(* IEC 61131-3 sources: JingjiangArm/moonboxpro_arm_8.4/Application/Application/任务列表/Main_Task/套色调整/套色新算法/PID_GET/Arc_pidh, 3 files *)

(* ---- DOUBLE_INTER.st ---- *)
(*@CES
Name=DOUBLE_INTER
Type=FunctionBlock
TypeGuid=6f9dac99-8de1-4efc-8465-68ac443b7d08
Guid=ffc9ca76-f385-4e76-b007-d8ddf6459d90
HasDeclaration=True
HasImplementation=True
*)
{DECLARATION}
FUNCTION DOUBLE_INTER : LREAL
VAR_INPUT
    (* --- 运行时输入 --- *)
    lrV_m_min   : LREAL;    (* 线速度 (m/min)，需在内部转换为 m/s *)
    lrY_Meas    : LREAL;    (* 测量套色误差 (mm) *)
    bEnable     : BOOL;     (* 控制器使能 *)

    (* --- 配置参数 (PSO 辨识与机械参数) --- *)
    lrPM_deg    : LREAL;    (* 目标相位裕度 (°) *)
    lrWc_Ts     : LREAL;    (* 归一化穿越频率 *)

    lrL         : LREAL;    (* 等效传输路径长度 (m) *)
    lrK_M       : LREAL;    (* 被控对象静态增益 (mm/deg) *)
    lrNK1       : LREAL;    (* 延迟物理量 *)
    lrC_SP      : LREAL;    (* 版辊等效周长 (m) *)

    (* --- 内部状态持久化指针 (外部传入) --- *)
    parrE       : POINTER TO ARRAY[1..2] OF LREAL; (* e(k-1), e(k-2) *)
    parrU       : POINTER TO ARRAY[1..2] OF LREAL; (* u(k-1), u(k-2) *)
END_VAR

VAR
    lrV_ms      : LREAL;    (* 转换后的线速度 m/s *)
    lrE_k       : LREAL;    (* 当前拍偏差 *)
    lrU_k       : LREAL;    (* 当前拍输出 *)

    lrTs        : LREAL;    (* 采样周期 *)
    lrA         : LREAL;    (* 极点 *)
    lrTau       : LREAL;    (* 传输延迟 *)
    lrPM_rad    : LREAL;    (* 相位裕度 (弧度) *)

    lrWc        : LREAL;    (* 穿越频率 *)
    lrWc_delay  : LREAL;    (* 受延迟约束的穿越频率上限 *)

    lrP_v       : LREAL;    (* 自适应极点 *)
    lrKc        : LREAL;    (* 自适应增益 *)

    lrAlpha     : LREAL;    (* Tustin 参数 2/Ts *)
    lrAlpha2    : LREAL;    (* Alpha 的平方 *)

    lrB0        : LREAL;    (* 差分方程系数 b0 *)
    lrB1        : LREAL;    (* 差分方程系数 b1 *)
    lrB2        : LREAL;    (* 差分方程系数 b2 *)

	//
	lrPi:LREAL:=3.14159265358979323846;
END_VAR
{IMPLEMENTATION}

(* ==========================================
   0. 空指针保护
   ========================================== *)
IF parrE = 0 OR parrU = 0 THEN
    DOUBLE_INTER := 0.0;
    RETURN;
END_IF;

(* ==========================================
   1. 单位转换与使能/速度保护
   ========================================== *)
lrV_ms := lrV_m_min / 60.0;(*单位对齐至m/s*)
IF lrC_SP<>0 THEN
	lrK_M := lrK_M * 36 / lrC_SP ;(*增益转换，从deg/mm转换到0.1丝/丝*)
ELSE
	lrK_M := 0.2;
END_IF
lrC_SP := lrC_SP / 1000.0 ;(*单位对齐至m*)

IF NOT bEnable THEN
    (* 未使能时，强制清空历史数组 *)
    parrE^[1] := 0.0;
    parrE^[2] := 0.0;
    parrU^[1] := 0.0;
    parrU^[2] := 0.0;
    DOUBLE_INTER := 0.0;
    RETURN;
END_IF;

IF lrV_ms < 0.1 THEN
    (* 速度过低保护，防止除零故障 *)
    DOUBLE_INTER := 0.0;
    RETURN;
END_IF;

(* ==========================================
   2. 计算物理模型参数与约束限制
   ========================================== *)
IF lrV_ms<>0 THEN
	lrTs  := lrC_SP / lrV_ms;
ELSE
	lrTs := 1;
END_IF

IF lrL<>0 THEN
	lrA   := lrV_ms / lrL;
ELSE
	lrA := 4.5;
END_IF
IF lrV_ms<>0 THEN
	lrTau := MAX(0.0, lrNK1 / lrV_ms);
ELSE
	lrTau := 0.6;
END_IF
lrPM_rad := lrPM_deg * lrPi / 180.0;

lrWc := lrWc_Ts / lrTs;
lrWc_delay := (lrPi / 2 - lrPM_rad) / MAX(lrTau, 0.001);

IF lrWc > lrWc_delay THEN
    lrWc := lrWc_delay;
END_IF;

(* ==========================================
   3. 反解自适应参数与 Tustin 离散化系数
   ========================================== *)
lrP_v := lrWc / TAN(lrPM_rad + (lrWc * lrTau));
lrKc  := (lrWc * lrWc) / (lrK_M * lrA * SQRT((lrWc * lrWc) + (lrP_v * lrP_v)));

lrAlpha  := 2.0 / lrTs;
lrAlpha2 := lrAlpha * lrAlpha;

lrB0 := lrKc * (lrAlpha + lrA) * (lrAlpha + lrP_v) / lrAlpha2;
lrB1 := lrKc * 2.0 * ((lrA * lrP_v) - lrAlpha2) / lrAlpha2;
lrB2 := lrKc * (lrA - lrAlpha) * (lrP_v - lrAlpha) / lrAlpha2;

(* ==========================================
   4. 差分方程执行
   ========================================== *)
lrE_k := lrY_Meas;

lrU_k := (lrB0 * lrE_k)
       + (lrB1 * parrE^[1])
       + (lrB2 * parrE^[2])
       + (2.0 * parrU^[1])
       - parrU^[2];

(* ==========================================
   5. 状态推移更新
   ========================================== *)
parrE^[2] := parrE^[1];
parrE^[1] := lrE_k;

parrU^[2] := parrU^[1];
parrU^[1] := lrU_k;

(* ==========================================
   6. 输出结果
   ========================================== *)
DOUBLE_INTER := lrU_k;

(* ---- Gc_PID_2024.st ---- *)
(*@CES
Name=Gc_PID_2024
Type=FunctionBlock
TypeGuid=6f9dac99-8de1-4efc-8465-68ac443b7d08
Guid=552ec7f6-cc2d-49c3-aeac-a3021bb272f5
HasDeclaration=True
HasImplementation=True
*)
{DECLARATION}
FUNCTION Gc_PID_2024 : REAL
(*2023.09.04.143809 增加加速积分环节*)
(*微调@2023.10.31.192825*)
(*2024.04.06.143012 增加pi的最大输出限值*)
(*2024.7.26.154629 将d值输出打开*)
(*2024.7.27.081735 输出超限了-从积分器里减*)
(*2024.9.12.174833*)
(*积分抗饱和增加注释@2025.1.13.171853*)
VAR_INPUT
	i_rTs:REAL;(*采样周期*)
	i_rP:REAL;
	i_rI:REAL;
	i_rD:REAL;
	i_rN:REAL;
	i_rU:REAL;(*控制器输入*)
	i_prYout: POINTER TO REAL;(*控制器输出*)

	i_parEk:POINTER TO ARRAY [1..2] OF REAL;(*误差寄存器 [e(k);e(k-1)]*)
	i_parYPk:POINTER TO ARRAY [1..2] OF REAL;(*比例控制输出寄存器*)
	i_parYIk:POINTER TO ARRAY [1..2] OF REAL;(*积分控制输出寄存器*)
	i_parYDk:POINTER TO ARRAY [1..2] OF REAL;(*微分控制输出寄存器*)
	i_parYPIDk:POINTER TO ARRAY [1..2] OF REAL;(*PID控制器输出寄存器*)
	(*2024.04.06.135400|增加了调整量的输出限值*)
	i_iMaxYPID:INT;(*最大的pid输出@增量*)
	i_iErrLimit_P:INT;(*Kp的误差限幅@2024.8.1.152553+*)
	i_iErrLimit_I:INT;(*积分的误差限幅@2024.8.1.152553+*)
END_VAR

VAR
	rP:REAL:=20.0;
	rI:REAL:=8.0;
	rD:REAL:=0;
	rN:REAL:=0;
	rTs:REAL:=0;

	rA:REAL:=0;(*加速度*)
	rA_max: REAL:=1.5;(*测试状态下写为定值*)

	rP2:REAL:=1.0;
	rI2:REAL:=0.5;(*用来控制那种加速补偿方式|=1 加速度补偿系数|=2 delta速度补偿方式*)
	rI2_A:REAL:=0.5;
	rPID_Y:REAL:=0;
	(*积分分离*)
	rE_max:REAL:=60.0;(*3*20*)
	rP_max:REAL:=40.0;(*2*rP*)

	(*加速补偿积分使用速度差系数2023.9.18*)
	rV0:REAL:=30.0;(*开始升速的速度*)(*测试状态下写为定值*)
	rVmax:REAL:=200.0;(*升速目标速度*)(*测试状态下写为定值*)
	rI2_v:REAL:=0;
	rDelta_V:REAL:=0;
	rEk_P: REAL;
	rEk_I: REAL;
	rDelta: REAL;
END_VAR
{IMPLEMENTATION}
rTs:=i_rTs;

rP:=i_rP;
rI:=i_rI;
rD:=i_rD;
rN:=i_rN;

(*先按照d不等于0的时候rN=1*)
IF rD=0 THEN
	rN:=0;
ELSE
	rN:=1;
END_IF

(*差分计算*)
i_parEk^[1]:=i_rU;
(*比例*)
(*2024.04.08.110035*)
(*i_prYPk^:=rP*i_parEk^[1];*)

(*对kp的误差值限幅@2024.8.1.152800*)
rEk_P:=i_parEk^[1];
IF i_iErrLimit_P<>0 THEN
	IF ABS(i_parEk^[1])>i_iErrLimit_P THEN
		rEk_P:=INT_TO_REAL(i_iErrLimit_P)*i_parEk^[1]/ABS(i_parEk^[1]);
	END_IF
END_IF
i_parYPk^[1]:=rP*rEk_P(*i_parEk^[1]*);
(*积分*)
(*积分的误差值限幅@2024.8.1.152800*)
rEk_I:=i_parEk^[2];
IF i_iErrLimit_I<>0 THEN
	IF ABS(i_parEk^[2])>i_iErrLimit_I THEN
		rEk_I:=INT_TO_REAL(i_iErrLimit_I)*i_parEk^[2]/ABS(i_parEk^[2]);
	END_IF
END_IF

i_parYIk^[1]:=i_parYIk^[2]+rI*rTs*rEk_I(*i_parEk^[2])*);
(*微分*)
i_parYDk^[1]:=i_parYDk^[2]*(1.0-rN*rTs)+rD*rN*(i_parEk^[1]-i_parEk^[2]);

(*2024.04.06.143033 先取消d值的使用吧*)
(*2024.7.26.141434  又把d值打开了*)
(*2024.04.08.110121*)
(*i_parYPIDk^[1]:=i_prYPk^+i_parYIk^[1]+i_parYDk^[1]*0;(*上面pi的输出*)*)
i_parYPIDk^[1]:=i_parYPk^[1]+i_parYIk^[1]+i_parYDk^[1];(*上面pi的输出*)

(*增加了限值输出@输出的变化量|2024.04.06.140853*)
rDelta:=ABS(i_parYPIDk^[1]-i_parYPIDk^[2]);

IF i_iMaxYPID<>0 THEN
	IF rDelta>i_iMaxYPID THEN(*输出超过了最大允许的变化量|做限值处理*)
		(*限值后的输出*)

		IF i_parYPIDk^[1]>i_parYPIDk^[2] THEN
			i_parYPIDk^[1]:=i_parYPIDk^[2]+i_iMaxYPID;
			(*从积分器里剔除@2024.7.27.081256*)
			i_parYIk^[1]:=i_parYIk^[1]-i_iMaxYPID;(*这种方式相当于是按照绝对位置输出@输出多少量,就减小多少*)
(*			i_parYIk^[1]:=i_parYIk^[1]-(rDelta-i_iMaxYPID);*)(*这种方式相当于是按照最大增量输出后不再输出*)

		ELSE
			i_parYPIDk^[1]:=i_parYPIDk^[2]-i_iMaxYPID;
			(*从积分器里剔除@2024.7.27.081256*)
			i_parYIk^[1]:=i_parYIk^[1]+i_iMaxYPID;(*这种方式相当于是按照绝对位置输出@输出多少量,就减小多少*)
(*			i_parYIk^[1]:=i_parYIk^[1]+(rDelta-i_iMaxYPID);*)(*这种方式相当于是按照最大增量输出后不再输出*)
		END_IF
(*
		IF ABS(i_parYPk^[1]-i_parYPk^[2])>=i_iMaxYPID THEN(*因为kp超过的,此时进行积分隔离@取消积分的叠加*)
			i_parYIk^[1]:=i_parYIk^[2];(*当前积分寄存器中的值和上一拍保持一致*)
		ELSE(*还有一部分积分起作用，超过限制值@只保留输出的积分部分*)
			i_parYIk^[1]:=i_parYPIDk^[1]-i_parYPk^[1];(*当前积分寄存器中的值和上一拍保持一致*)
		END_IF
*)
	END_IF
ELSE;(*保持之前的*)
END_IF

(*更新寄存器的值-注意顺序*)
i_parEk^[2]:=i_parEk^[1];
i_parYPk^[2]:=i_parYPk^[1];(*2024.04.08.110707+*)
i_parYIk^[2]:=i_parYIk^[1];
i_parYDk^[2]:=i_parYDk^[1];
i_parYPIDk^[2]:=i_parYPIDk^[1];

i_prYout^:=i_parYPIDk^[1];

(* ---- Gc_PID_2025.st ---- *)
(*@CES
Name=Gc_PID_2025
Type=FunctionBlock
TypeGuid=6f9dac99-8de1-4efc-8465-68ac443b7d08
Guid=460d2dc5-80dd-4599-9edb-64334fe92a43
HasDeclaration=True
HasImplementation=True
*)
{DECLARATION}
FUNCTION Gc_PID_2025 : REAL
(*2025.1.15.095113@增加误差阈值,超过该值按照最大值输出。范围内按照pi控制器输出*)
VAR_INPUT
	i_rTs:REAL;(*采样周期*)
	i_rP:REAL;
	i_rI:REAL;
	i_rD:REAL;
	i_rN:REAL;
	i_rU:REAL;(*控制器输入*)
	i_prYout: POINTER TO REAL;(*控制器输出*)

	i_parEk:POINTER TO ARRAY [1..2] OF REAL;(*误差寄存器 [e(k);e(k-1)]*)
	i_parYPk:POINTER TO ARRAY [1..2] OF REAL;(*比例控制输出寄存器*)
	i_parYIk:POINTER TO ARRAY [1..2] OF REAL;(*积分控制输出寄存器*)
	i_parYDk:POINTER TO ARRAY [1..2] OF REAL;(*微分控制输出寄存器*)
	i_parYPIDk:POINTER TO ARRAY [1..2] OF REAL;(*PID控制器输出寄存器*)
END_VAR

VAR
	rP:REAL:=20.0;
	rI:REAL:=8.0;
	rD:REAL:=0;
	rN:REAL:=0;
	rTs:REAL:=0;
END_VAR
{IMPLEMENTATION}
rTs:=i_rTs;

rP:=i_rP;
rI:=i_rI;
rD:=i_rD;
rN:=i_rN;

(*先按照d不等于0的时候rN=1*)
IF rD=0 THEN
	rN:=0;
ELSE
	rN:=1;
END_IF

(*差分计算*)
i_parEk^[1]:=i_rU;

(*超过阈值按照最大值输出*)
(*比例*)
i_parYPk^[1]:=rP*i_parEk^[1];
(*积分*)
i_parYIk^[1]:=i_parYIk^[2]+rI*rTs*i_parEk^[2];
(*微分*)
i_parYDk^[1]:=i_parYDk^[2]*(1.0-rN*rTs)+rD*rN*(i_parEk^[1]-i_parEk^[2]);
(*总输出*)
i_parYPIDk^[1]:=i_parYPk^[1]+i_parYIk^[1]+i_parYDk^[1];(*上面pi的输出*)

(*更新寄存器的值-注意顺序*)
i_parEk^[2]:=i_parEk^[1];
i_parYPk^[2]:=i_parYPk^[1];(*2024.04.08.110707+*)
i_parYIk^[2]:=i_parYIk^[1];
i_parYDk^[2]:=i_parYDk^[1];
i_parYPIDk^[2]:=i_parYPIDk^[1];

i_prYout^:=i_parYPIDk^[1];
